FUNCTION_BLOCK FB_EtherCATFrameDiag_1
VAR_INPUT
	wFrmXWcState 		: WORD;
	wReqZeroMask 		: WORD := 16#FFFF; (* bit TRUE: require wFrmXWcState.bit = FALSE, bit FALSE: ignore wFrmXWcState.bit *)
END_VAR
VAR_OUTPUT
	bFrameWcStateOK		: BOOL;
END_VAR
VAR
END_VAR

(* set/clear frame flag *)
bFrameWcStateOK := ((wFrmXWcState AND wReqZeroMask) = 0);

END_FUNCTION_BLOCK

(* stored: Version 1.1.0.1, ProductVersion 3.1.4024.15
   POU FB_EtherCATFrameDiag_1: Id {b3e3f95f-0d61-40b2-a345-7abaa0246d82}, SpecialFunc None *)
